// TIA Portal project "Project8" (V19)

(* hardware
DEVICE "S7-1500/ET200MP station_1"  S7-1500 station
   slot 0: "Rail_0"  Rack  6ES7 590-1***0-0AA0
   slot 1: "PLC_1"  CPU 1511-1 PN  6ES7 511-1AK01-0AB0  V2.9
      slot 3: "CPU display_1"  6ES7591-1AA00-0AA0
      slot 32768: "PROFINET interface_1"  X1
         slot 32769: "Port_1"  X1 P1
         slot 32770: "Port_2"  X1 P2
      slot 34817: "Virtual CP interface port_1"  Virtual CP interface port  Virtual CP interface port
   slot 2: "DI 16x24VDC / DQ 16x24VDC/0.5A BA_1"  DI 16x24VDC/DQ 16x24VDC/0.5A BA  6ES7 523-1BL00-0AA0  V1.1
*)

// ===== PLC "PLC_1"  CPU 1511-1 PN =====

VAR_GLOBAL   // PLC tag table "Default tag table"
   "Tag_1" AT %I0.0 : Bool;
   "Tag_2" AT %I0.1 : Bool;
   "Tag_3" AT %Q0.1 : Bool;
END_VAR

DATA_BLOCK "Data_block_1"   // DB1
{ S7_Optimized_Access := 'FALSE' }
VERSION : 0.1
   VAR
      I_Start : Bool;
      I_Stop : Bool;
      Q_Lamp : Bool;
   END_VAR
BEGIN
END_DATA_BLOCK

DATA_BLOCK "DB_Tank"   // DB2
{ S7_Optimized_Access := 'FALSE' }
VERSION : 0.1
   VAR
      Was_Running : Bool;
      V_Out_Saved : Real;
      SP_Level : Real := 50.0;
      V_In : Real;
      V_Out : Real;
      L_Level : Real;
   END_VAR
BEGIN
END_DATA_BLOCK

ORGANIZATION_BLOCK "Main"   // OB1, LAD, ProgramCycle
TITLE = "Main Program Sweep (Cycle)"
{ S7_Optimized_Access := 'TRUE' }
VERSION : 0.1
   VAR_INPUT
      Initial_Call : Bool;   // Initial call of this OB
      Remanence : Bool;   // =True, if remanent data are available
   END_VAR
BEGIN

REGION Network 1
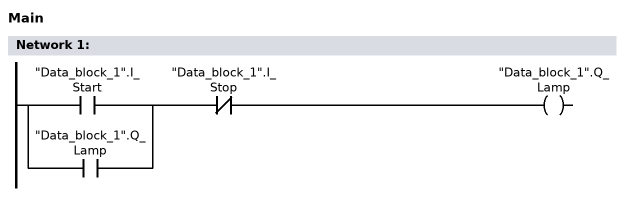
   RUNG wire#powerrail
      Contact( "Data_block_1".I_Start )
      wire#w1
      I_Contact( "Data_block_1".I_Stop )
      Coil( "Data_block_1".Q_Lamp )
   END_RUNG
   RUNG wire#powerrail
      Contact( "Data_block_1".Q_Lamp )
   END_RUNG wire#w1
   // the same network as SCL:
   "Data_block_1".Q_Lamp := ("Data_block_1".I_Start OR "Data_block_1".Q_Lamp) AND NOT "Data_block_1".I_Stop;
END_REGION
END_ORGANIZATION_BLOCK

ORGANIZATION_BLOCK "OB_PID_Level"   // OB30, SCL, CyclicInterrupt
{ S7_Optimized_Access := 'TRUE' }
VERSION : 0.1
   VAR_INPUT
      Initial_Call : Bool;   // Initial call of this OB
      Event_Count : Int;   // Events discarded
   END_VAR
BEGIN
   "PID_Level"(Setpoint := "DB_Tank".SP_Level,
               Input := "DB_Tank".L_Level,
               Output => "DB_Tank".V_In);

   IF "Data_block_1".Q_Lamp AND NOT "DB_Tank".Was_Running THEN
       "DB_Tank".V_Out := "DB_Tank".V_Out_Saved;
   ELSIF NOT "Data_block_1".Q_Lamp AND "DB_Tank".Was_Running THEN
       "DB_Tank".V_Out_Saved := "DB_Tank".V_Out;
   END_IF;

   IF NOT "Data_block_1".Q_Lamp THEN
       "DB_Tank".V_In := 0.0;
       "DB_Tank".V_Out := 0.0;
   END_IF;

   "DB_Tank".Was_Running := "Data_block_1".Q_Lamp;
   IF NOT "Data_block_1".Q_Lamp THEN
       "DB_Tank".V_In := 0.0;
       "DB_Tank".V_Out := 0.0;
   END_IF;

   "DB_Tank".Was_Running := "Data_block_1".Q_Lamp;
END_ORGANIZATION_BLOCK